// TIA Portal V21 export
// export: Created 2026-08-21T20:18:50.7711144Z, ExportSetting None, DisplayName Totally Integrated Automation Portal, DisplayVersion V21, DisplayName STEP 7 Professional, DisplayVersion V21, DisplayName STEP 7 Safety, DisplayVersion V21, DisplayName Tech WebApplication, DisplayVersion V21, DisplayName WinCC Basic/Comfort/Advanced, DisplayVersion V21, DisplayName WinCC Professional, DisplayVersion V21, DisplayName WinCC Unified, DisplayVersion V21
FUNCTION "FIC100" : Void   // FC5, FBD
{ S7_Optimized_Access := 'TRUE' }
// stored: SetENOAutomatically false
   VAR_TEMP
      Temp : "DigVal";
      State : "Service_States";
      Interlock : "DigVal";
   END_VAR
BEGIN

REGION Network 1: PIDConL interconnections
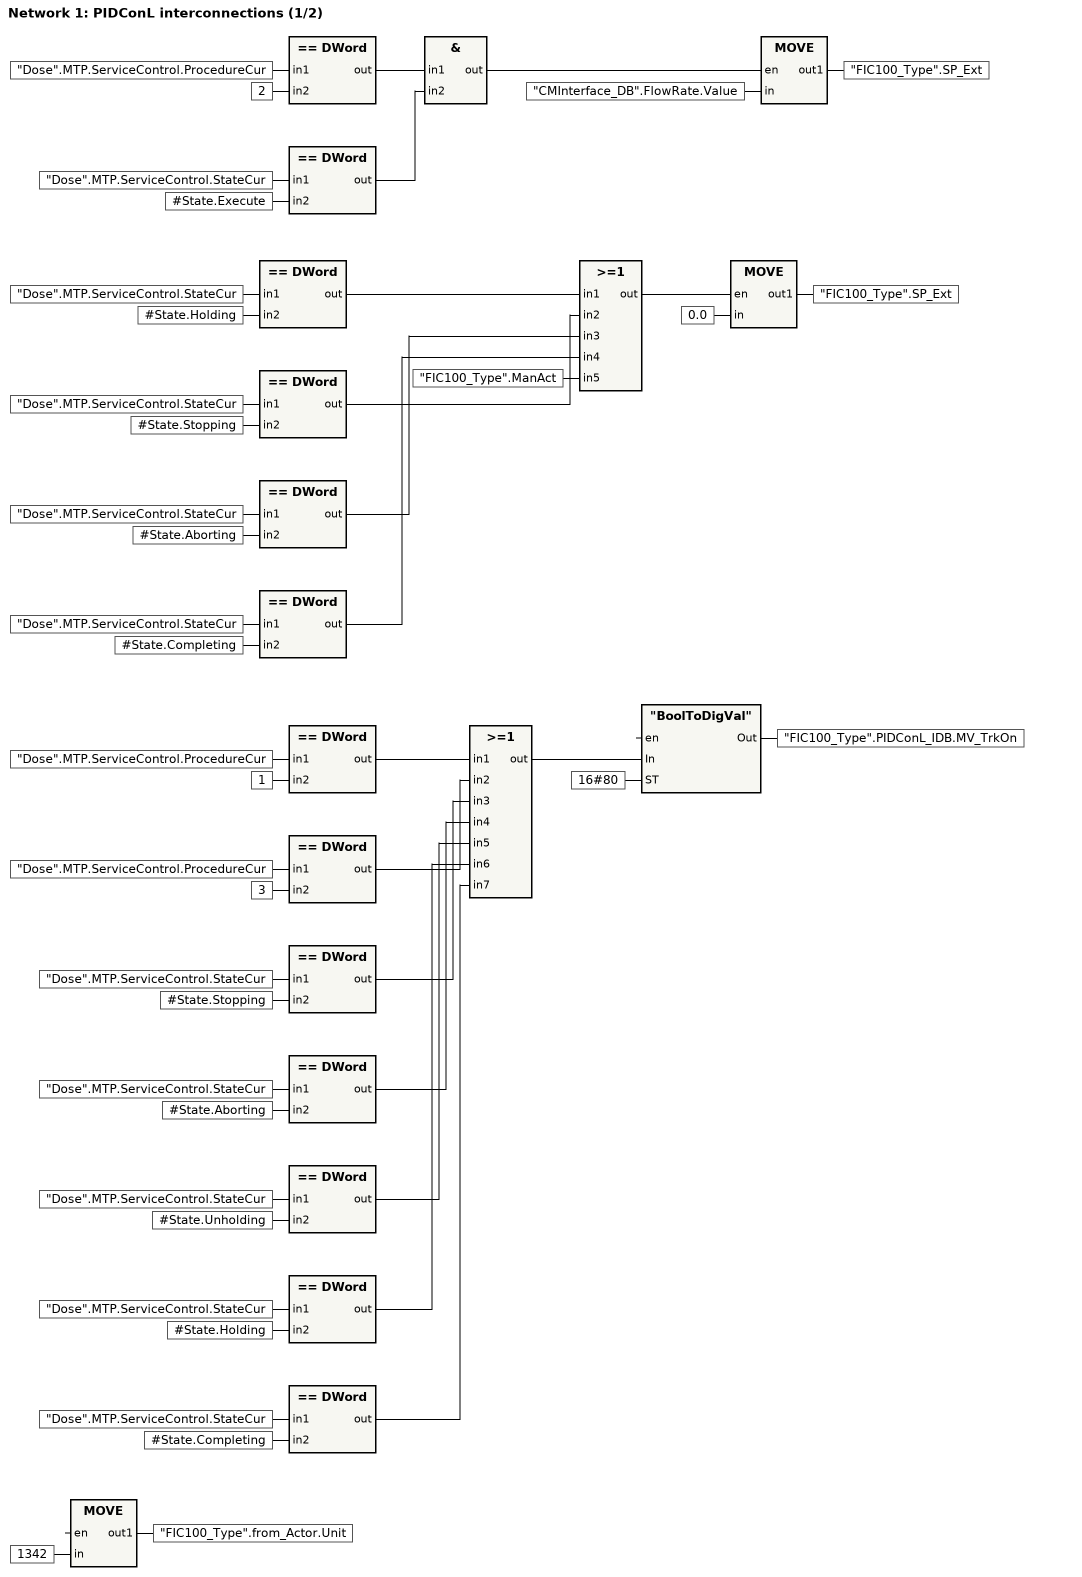
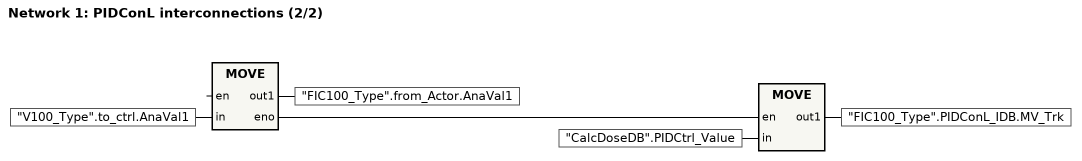
   IF ("Dose".MTP.ServiceControl.ProcedureCur = 2) AND ("Dose".MTP.ServiceControl.StateCur = #State.Execute) THEN
       "FIC100_Type".SP_Ext := "CMInterface_DB".FlowRate.Value;
   END_IF;
   IF ("Dose".MTP.ServiceControl.StateCur = #State.Holding) OR ("Dose".MTP.ServiceControl.StateCur = #State.Stopping) OR ("Dose".MTP.ServiceControl.StateCur = #State.Aborting) OR ("Dose".MTP.ServiceControl.StateCur = #State.Completing) OR "FIC100_Type".ManAct THEN
       "FIC100_Type".SP_Ext := 0.0;
   END_IF;
   "BoolToDigVal"(In := ("Dose".MTP.ServiceControl.ProcedureCur = 1) OR ("Dose".MTP.ServiceControl.ProcedureCur = 3) OR ("Dose".MTP.ServiceControl.StateCur = #State.Stopping) OR ("Dose".MTP.ServiceControl.StateCur = #State.Aborting) OR ("Dose".MTP.ServiceControl.StateCur = #State.Unholding) OR ("Dose".MTP.ServiceControl.StateCur = #State.Holding) OR ("Dose".MTP.ServiceControl.StateCur = #State.Completing),
                  ST := 16#80,
                  Out => "FIC100_Type".PIDConL_IDB.MV_TrkOn);
   "FIC100_Type".from_Actor.Unit := 1342;
   "FIC100_Type".from_Actor.AnaVal1 := "V100_Type".to_ctrl.AnaVal1;
   "FIC100_Type".PIDConL_IDB.MV_Trk := "CalcDoseDB".PIDCtrl_Value;
END_REGION

REGION Network 2: PIDCon
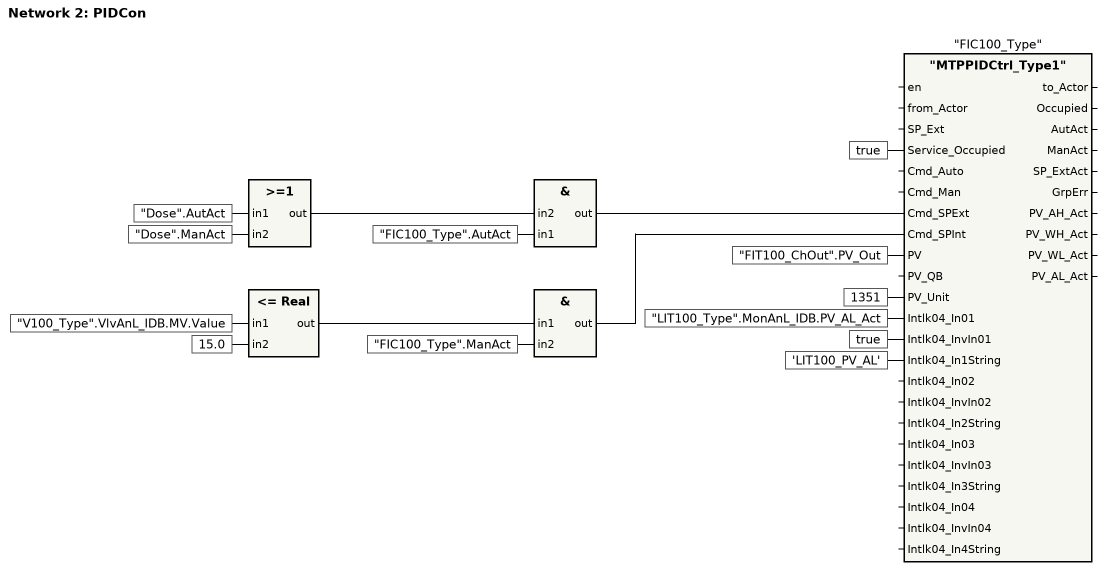
   "FIC100_Type"(Service_Occupied := true,   // "MTPPIDCtrl_Type1"
                 Cmd_SPExt := ("Dose".AutAct OR "Dose".ManAct) AND "FIC100_Type".AutAct,
                 Cmd_SPInt := ("V100_Type".VlvAnL_IDB.MV.Value <= 15.0) AND "FIC100_Type".ManAct,
                 PV := "FIT100_ChOut".PV_Out,
                 PV_Unit := 1351,
                 Intlk04_In01 := "LIT100_Type".MonAnL_IDB.PV_AL_Act,
                 Intlk04_InvIn01 := true,
                 Intlk04_In1String := 'LIT100_PV_AL');
END_REGION
END_FUNCTION
